// TIA Portal V20 export
// export: Created 2026-10-20T18:55:04.8717817Z, ExportSetting None, DisplayName Totally Integrated Automation Portal, DisplayVersion V20 Update 6, DisplayName TIA Portal Openness, DisplayVersion V20 Update 6, DisplayName TIA Portal Version Control Interface, DisplayVersion V20 Update 6, DisplayName SINAMICS Startdrive Advanced, DisplayVersion V20 SP1, DisplayName SINAMICS Startdrive G130, G150, S120, S150, SINAMICS MV, G220, S200, S210, DisplayVersion V20 SP1, DisplayName SINAMICS Startdrive G110M, G120, G120C, G120D, G120P, G115D, DisplayVersion V20 SP1, DisplayName STEP 7 Professional, DisplayVersion V20 Update 6, DisplayName STEP 7 Safety, DisplayVersion V20 Update 2, DisplayName WinCC Basic/Comfort/Advanced, DisplayVersion V20 Update 6, DisplayName WinCC Unified, DisplayVersion V20 Update 6
VAR_GLOBAL   // PLC tag table "IO_VFDs_3"
   C3101_MainSetpoint AT %QW858 : Word;
   C3101_StatusWord AT %IW2426 : Word;
   C3206_ActualSpeed AT %IW2584 : Word;
   VTD3_MainSetpoint AT %QW496 : Word;
   C3103_StatusWord AT %IW2450 : Word;
   C3108_ControlWord AT %QW956 : Word;
   C3106_MainSetpoint AT %QW878 : Word;
   C3208_ControlWord AT %QW988 : Word;
   C3103_ControlWord AT %QW864 : Word;
   C3207_ActualCurrent AT %IW2598 : Word;
   C3105_ActualCurrent AT %IW2478 : Word;
   C3202_ActualCurrent AT %IW2538 : Word;
   C3204_ActualCurrent AT %IW2562 : Word;
   C3108_MainSetpoint AT %QW958 : Word;
   C3108_ActualSpeed AT %IW2512 : Word;
   C3208_MainSetpoint AT %QW990 : Word;
   C3205_ActualSpeed AT %IW2572 : Word;
   C3207_MainSetpoint AT %QW986 : Word;
   C3101_ActualCurrent AT %IW2430 : Word;
   VTD3_ControlWord AT %QW494 : Word;
   C3106_ControlWord AT %QW876 : Word;
   C3203_MainSetpoint AT %QW970 : Word;
   C3208_ActualCurrent AT %IW2610 : Word;
   C3102_ActualCurrent AT %IW2442 : Word;
   C3105_ControlWord AT %QW872 : Word;
   CVTD3_MainSetpoint AT %QW536 : Word;
   CVTD3_StatusWord AT %IW2414 : Word;
   C3202_ControlWord AT %QW964 : Word;
   VTD3_ActualSpeed AT %IW1034 : Word;
   C3103_ActualCurrent AT %IW2454 : Word;
   C3105_StatusWord AT %IW2474 : Word;
   C3201_ActualCurrent AT %IW2526 : Word;
   C3203_ControlWord AT %QW968 : Word;
   C3106_StatusWord AT %IW2486 : Word;
   C3205_MainSetpoint AT %QW978 : Word;
   C3104_ControlWord AT %QW868 : Word;
   CVTD3_ActualCurrent AT %IW2418 : Word;
   C3201_MainSetpoint AT %QW962 : Word;
   C3102_MainSetpoint AT %QW862 : Word;
   C3203_StatusWord AT %IW2546 : Word;
   VTD3_ActualCurrent AT %IW1036 : Word;
   C3102_StatusWord AT %IW2438 : Word;
   C3205_StatusWord AT %IW2570 : Word;
   C3207_StatusWord AT %IW2594 : Word;
   C3103_ActualSpeed AT %IW2452 : Word;
   C3207_ControlWord AT %QW984 : Word;
   CVTD3_ActualSpeed AT %IW2416 : Word;
   C3104_ActualSpeed AT %IW2464 : Word;
   C3104_ActualCurrent AT %IW2466 : Word;
   C3201_ControlWord AT %QW960 : Word;
   C3204_ActualSpeed AT %IW2560 : Word;
   C3208_ActualSpeed AT %IW2608 : Word;
   C3106_ActualCurrent AT %IW2490 : Word;
   C3105_ActualSpeed AT %IW2476 : Word;
   C3208_StatusWord AT %IW2606 : Word;
   C3203_ActualSpeed AT %IW2548 : Word;
   C3205_ControlWord AT %QW976 : Word;
   C3206_ActualCurrent AT %IW2586 : Word;
   C3206_MainSetpoint AT %QW982 : Word;
   C3108_StatusWord AT %IW2510 : Word;
   C3101_ActualSpeed AT %IW2428 : Word;
   C3201_ActualSpeed AT %IW2524 : Word;
   C3108_ActualCurrent AT %IW2514 : Word;
   C3203_ActualCurrent AT %IW2550 : Word;
   C3201_StatusWord AT %IW2522 : Word;
   C3204_ControlWord AT %QW972 : Word;
   C3202_MainSetpoint AT %QW966 : Word;
   C3104_MainSetpoint AT %QW870 : Word;
   C3206_StatusWord AT %IW2582 : Word;
   C3207_ActualSpeed AT %IW2596 : Word;
   C3204_MainSetpoint AT %QW974 : Word;
   C3204_StatusWord AT %IW2558 : Word;
   CVTD3_ControlWord AT %QW534 : Word;
   C3107_StatusWord AT %IW2498 : Word;
   C3102_ControlWord AT %QW860 : Word;
   VTD3_StatusWord AT %IW1032 : Word;
   C3206_ControlWord AT %QW980 : Word;
   C3102_ActualSpeed AT %IW2440 : Word;
   C3202_ActualSpeed AT %IW2536 : Word;
   C3103_MainSetpoint AT %QW866 : Word;
   C3205_ActualCurrent AT %IW2574 : Word;
   C3101_ControlWord AT %QW856 : Word;
   C3105_MainSetpoint AT %QW874 : Word;
   C3107_ControlWord AT %QW952 : Word;
   C3107_ActualSpeed AT %IW2500 : Word;
   C3107_ActualCurrent AT %IW2502 : Word;
   C3104_StatusWord AT %IW2462 : Word;
   C3202_StatusWord AT %IW2534 : Word;
   C3107_MainSetpoint AT %QW954 : Word;
   C3106_ActualSpeed AT %IW2488 : Word;
   C3107_ActualTorque AT %IW2504 : Word;
   VTD3_ActualTorque AT %IW1038 : Word;
   C3201_ActualTorque AT %IW2528 : Word;
   C3204_ActualTorque AT %IW2564 : Word;
   C3108_ActualTorque AT %IW2516 : Word;
   C3208_ActualTorque AT %IW2612 : Word;
   C3101_ActualTorque AT %IW2432 : Word;
   C3207_ActualTorque AT %IW2600 : Word;
   C3102_ActualTorque AT %IW2444 : Word;
   C3106_ActualTorque AT %IW2492 : Word;
   C3203_ActualTorque AT %IW2552 : Word;
   C3205_ActualTorque AT %IW2576 : Word;
   C3202_ActualTorque AT %IW2540 : Word;
   C3104_ActualTorque AT %IW2468 : Word;
   C3103_ActualTorque AT %IW2456 : Word;
   C3105_ActualTorque AT %IW2480 : Word;
   C3206_ActualTorque AT %IW2588 : Word;
   CVTD3_ActualTorque AT %IW2420 : Word;
   VTD3_AccFactor AT %QW1521 : Word;
END_VAR
